(* IEC 61131-3 sources: moqui-plc/codesys-v4/moqui-plc.fbsdev/moqui.iecapp^/moqui/framework/src/main/org/moqui/diagnostics, 2 files *)

(* ---- RemoteIoModuleDiagnostics.fb.st ---- *)
FUNCTION_BLOCK RemoteIoModuleDiagnostics

	VAR_INPUT
		moduleName : STRING;
	END_VAR
	VAR_OUTPUT
		error : BOOL;
		diagnosisInfo : STRING;
	END_VAR
	VAR
		byteArrayBuffer : ARRAY[0..1] OF BYTE;
		(* ABB parameters *)
		deviceState : BYTE;
		parameterState : BYTE;
	END_VAR

	error := TRUE;

	(*
	(* Example diagnostic code *)
	IF moduleName = 'io1' THEN
		toByteArray(inputWord := io1DeviceInformationBlock, byteArray => byteArrayBuffer);
		deviceState := byteArrayBuffer[0];
		parameterState := byteArrayBuffer[1];
	(*
	ELSIF moduleName = 'io2' THEN
		toByteArray(inputWord := io2DeviceInformationBlock, byteArray => byteArrayBuffer);
	    deviceState := byteArrayBuffer[0];
	    parameterState := byteArrayBuffer[1];
	*)
	ELSE
		RETURN;
	END_IF;

	(* The actual state of the remote IO module *)
	diagnosisInfo := concat(concat('IO module ', moduleName), ' diagnosis info: ');
	CASE deviceState OF
		0 : diagnosisInfo := concat('STATE_PREOP', diagnosisInfo);
		1 : diagnosisInfo := concat('STATE_OPERATION', diagnosisInfo);
		2 : diagnosisInfo := concat('STATE_ERROR', diagnosisInfo); RETURN;
		3 : diagnosisInfo := concat('STATE_IP_ERROR', diagnosisInfo); RETURN;
		4 : diagnosisInfo := concat('STATE_CYCLIC_OPERATION', diagnosisInfo);
	ELSE
		RETURN;
	END_CASE;

	CASE parameterState OF
		0 : diagnosisInfo := concat('PARA_STATE_NO_PARA', diagnosisInfo);
		1 : diagnosisInfo := concat('PARA_STATE_PARA_ACTIVE', diagnosisInfo);
		2 : diagnosisInfo := concat('PARA_STATE_PARA_DONE', diagnosisInfo);
		3 : diagnosisInfo := concat('PARA_STATE_PARA_DONE', diagnosisInfo);
		4 : diagnosisInfo := concat('PARA_STATE_ERROR', diagnosisInfo); RETURN;
	ELSE
		RETURN;
	END_CASE;

	(* etc. *)
	*)

	error := FALSE;
	END_FUNCTION_BLOCK

(* ---- SignalMgmt.fb.st ---- *)
(* Signal supervisor *)
FUNCTION_BLOCK SignalMgmt

	VAR_INPUT
		operationType : SignalMgmtOperatingMode;
		(* Signal metadata *)
	    code : WORD; (* Unique ID for assigning a static priority to signals of the same category *)
		category : SignalCategory; (* Signal type: Static category/priority level + reset policy *)
		resetPol : ResetPolicy := ResetPolicy.UnconditionedReset;
	    outputAction : SignalOutputAction := SignalOutputAction.None; (* Response output/action to the signal detection (e.g. ImmediateStop, EmergencyStop, etc.). *)
		(* Activation condition (condition of failure) or trigger policy for the signal, as a boolean expression *)
	    activationCondition : BOOL;
		(*
	     * Condition for auto conditioned reset for the signal, as a boolean expression (e.g. MachineNotRunning).
	     * The reset condition or policy is considered only if an activation policy has
	     * been selected during the configuration phase.
		 *)
		autoResetCondition : BOOL;
	    (* Reset commands *)
	    reset : BOOL; (* Unconditioned manual/external reset *)
	    auxReset : BOOL; (* Auxiliary key or command *)
	    (* Selective reset *)
	    selectiveResetTrigger : BOOL;
	    selectiveResetCode : WORD;
	    (* Logger name for recording events associated with signals *)
	    loggerName : STRING := '';
	END_VAR
	VAR_OUTPUT
	    cumulativeOutputAction : DWORD := SignalOutputAction.None; (* Cumulative output (stop) for the current cycle *)
	    activeCategory : SignalCategory; (* Most severe category active *)
	    (* Reset availability indicators (updated each cycle in Prepare+Process, for operator feedback) *)
	    resetEnable : BOOL; (* TRUE if at least one active signal has cause gone and requires manual reset *)
	    auxResetEnable : BOOL; (* TRUE if at least one active signal has cause gone and accepts aux reset *)
		(* Invalid signal code or missing loggerName; kept until the next Reset *)
		error : BOOL := FALSE;
	END_VAR
	VAR
		(* Logger facade *)
	    logger : LoggerFacade;
	    (* Persistent signal log *)
	    signalList : ARRAY[1..MoquiConf.SIGNAL_LIST_MAX_SIZE] OF BOOL;
	    (* Variables for detecting reset edges *)
	    resetOld : BOOL;
	    resetActivation : BOOL;
	    auxResetOld : BOOL;
	    auxResetActivation : BOOL;
	    selectiveResetOld : BOOL;
	    selectiveResetActivation : BOOL;
	    requiresManualReset : BOOL;
		(* Cumulative output of the previous cycle, so that it is logged on change only *)
		cumulativeOutputActionOld : DWORD := SignalOutputAction.None;
		i : UINT;
	END_VAR

	(* Args validation *)
	IF (loggerName = '') THEN error := TRUE; RETURN; END_IF;

	(* Logger facade init *)
	logger.enable := TRUE; logger.loggerName := loggerName;

	CASE operationType OF
	    SignalMgmtOperatingMode.Reset :
			logger(message := 'Signal management reset.', level := LogLevel.DEBUG);
	        error := FALSE;
	        cumulativeOutputActionOld := SignalOutputAction.None;
	        FOR i := 1 TO MoquiConf.SIGNAL_LIST_MAX_SIZE DO signalList[i] := FALSE; END_FOR;
	        resetOld := FALSE; auxResetOld := FALSE; selectiveResetOld := FALSE;
	        cumulativeOutputAction := SignalOutputAction.None;
	        activeCategory := SignalCategory.Information;
	        resetEnable := FALSE; auxResetEnable := FALSE;

	    SignalMgmtOperatingMode.Prepare :
	        (* The previous cycle is complete: log its cumulative output if it changed *)
	        IF cumulativeOutputAction <> cumulativeOutputActionOld THEN
	            logger(message := concat('Signal cumulative output: ', DWORD_TO_STRING(cumulativeOutputAction)), level := LogLevel.Info);
	            cumulativeOutputActionOld := cumulativeOutputAction;
	        END_IF;
	        (* Detection of reset edges valid for the entire cycle  *)
	        resetActivation := reset AND NOT resetOld;
	        resetOld := reset;
	        auxResetActivation := auxReset AND NOT auxResetOld;
	        auxResetOld := auxReset;
	        selectiveResetActivation := selectiveResetTrigger AND NOT selectiveResetOld;
	        selectiveResetOld := selectiveResetTrigger;
	        (* Init for the current cycle *)
	        cumulativeOutputAction := SignalOutputAction.None;
	        activeCategory := SignalCategory.Information;
	        resetEnable := FALSE; auxResetEnable := FALSE;

	    SignalMgmtOperatingMode.Process :
	        (* Bounds check *)
	        IF (code < 1) OR (code > MoquiConf.SIGNAL_LIST_MAX_SIZE) THEN
	            IF NOT error THEN logger(message := concat('Invalid signal code: ', WORD_TO_STRING(code)), level := LogLevel.Error); END_IF;
	            error := TRUE;
	            RETURN;
	        END_IF;

	        (*
	         * Determine if manual reset is required.
	         * - Alarm, Anomaly: require manual reset unless resetPol = AutoReset
	         * - Warning, Information: always auto-reset
	         *)
	        CASE category OF
	            SignalCategory.Alarm, SignalCategory.Anomaly:
	                (* Both require manual reset by default; AutoReset policy overrides this *)
	                requiresManualReset := (resetPol <> ResetPolicy.AutoReset);
	            SignalCategory.Warning, SignalCategory.Information:
	                requiresManualReset := FALSE;
	        END_CASE;

	        (* Check the activation condition *)
	        IF activationCondition AND NOT signalList[code] THEN
				signalList[code] := TRUE;
	            (* Trigger the logger *)
	            logger(enable := TRUE, loggerName := loggerName, level := LogLevel.Fatal,
					message := concat(concat('Signal code: ', WORD_TO_STRING(code)), ' active.'));
	        END_IF;

	        (*
	         * Reset logic.
	         * An active signal is reset if the physical cause has disappeared (NOT activationCondition)
	         * AND one of the following re-entry conditions occurs, filtered by resetPol:
	         *   - Auto-reset (Warning/Information, or Alarm/Anomaly with AutoReset policy)
	         *   - Unconditioned manual reset: always allowed for Alarm
	         *   - Aux reset: only if resetPol = AuxReset
	         *   - Conditioned reset: only if resetPol = AutoConditionedReset / AutoProvisionalReset / AutoPriorityReset
	         *   - Selective reset: always allowed (supervisor override)
	         *)
	        IF NOT activationCondition AND signalList[code] THEN
	            IF NOT requiresManualReset THEN
	                (* Auto-reset: Anomaly, Warning, Information, or Alarm with AutoReset policy *)
	                signalList[code] := FALSE;
	            ELSIF resetActivation THEN
	                (* Unconditioned manual reset *)
	                signalList[code] := FALSE;
	            ELSIF auxResetActivation AND (resetPol = ResetPolicy.AuxReset) THEN
	                (* Aux reset: only if explicitly configured *)
	                signalList[code] := FALSE;
	            ELSIF autoResetCondition AND (
	                    resetPol = ResetPolicy.AutoConditionedReset OR
	                    resetPol = ResetPolicy.AutoProvisionalReset OR
	                    resetPol = ResetPolicy.AutoPriorityReset) THEN
	                (* Conditioned reset: only if explicitly configured *)
	                signalList[code] := FALSE;
	            ELSIF selectiveResetActivation AND (selectiveResetCode = code) THEN
	                (* Selective reset from external supervision: always allowed *)
	                signalList[code] := FALSE;
	            END_IF;

	            IF NOT signalList[code] THEN
	                logger(message := concat(concat('Signal code: ', WORD_TO_STRING(code)), ' reset.'), level := LogLevel.Info);
	            END_IF;
	        END_IF;

	        (* Cumulative stop bitmask *)
	        IF signalList[code] THEN
	            cumulativeOutputAction := cumulativeOutputAction OR outputAction;

	            (* Track the most severe category active in this cycle *)
	            IF category < activeCategory THEN
	                activeCategory := category;
	            END_IF;
	        END_IF;

	        (* Reset availability: signal is active, cause is gone, manual reset is required *)
	        IF signalList[code] AND NOT activationCondition AND requiresManualReset THEN
	            resetEnable := TRUE;
	        END_IF;
	        IF signalList[code] AND NOT activationCondition AND (resetPol = ResetPolicy.AuxReset) THEN
	            auxResetEnable := TRUE;
	        END_IF;
	END_CASE;
	END_FUNCTION_BLOCK
